TYPE "ST_PartContext"
VERSION : 0.1
   STRUCT
      "Uid" : String[64];
      "Present" : Bool;
      "CarrierKind" : DInt;
      "Result" : "ST_PartResult";
      "Parents" : Array[1..8] of String[64];
   END_STRUCT;
END_TYPE
